FUNCTION_BLOCK fbShutterAct
VAR_INPUT
	Config :  stShutterConfig;
	OpenRelay : iRelay;
	CloseRelay : iRelay;
END_VAR
VAR_OUTPUT
	State : stShutterState;
END_VAR
VAR_IN_OUT

END_VAR
VAR
	CmdOpen : BOOL;
	CmdClose : BOOL;
	OutputCheckTimer : TON;
END_VAR

VAR CONSTANT
	OutputCheckCycleTime: TIME := T#50MS;
END_VAR
VAR RETAIN
	HeightTime: TIME := T#0S;
	AngleTime: TIME := T#0S;
END_VAR


// Both signals must not be set at the same time
IF CmdOpen AND CmdClose THEN
	CmdOpen := FALSE;
	CmdClose := FALSE;
END_IF

// Reset signal if shutter reached fully open position with overstep
IF CmdOpen AND HeightTime >= Config.HeightTravelTime + Config.HeightTravelTimeOverstep THEN
	CmdOpen := FALSE;
END_IF

// Reset signal if shutter reached fully close position
IF CmdClose AND HeightTime <= T#0S AND AngleTime <= T#0S THEN
	CmdClose := FALSE;
END_IF

// Write physical outputs and update shutter state
IF CmdOpen AND NOT CmdClose THEN
    CloseRelay.Reset();
    OpenRelay.Set();
	State.StateType := eShutterStateType.OPENING;
ELSIF CmdClose AND NOT CmdOpen THEN
    OpenRelay.Reset();
    CloseRelay.Set();
	State.StateType := eShutterStateType.CLOSING;
ELSE
    OpenRelay.Reset();
    CloseRelay.Reset();
	State.StateType := eShutterStateType.IDLE;
END_IF

// Count time and accumulate when signals are set
OutputCheckTimer(IN := CmdOpen OR CmdClose, PT := OutputCheckCycleTime);
IF OutputCheckTimer.Q THEN
	IF CmdOpen THEN
		// Open fins first before moving up
		IF AngleTime < Config.AngleTravelTime THEN
			AngleTime := AngleTime + OutputCheckCycleTime;
		ELSIF HeightTime < Config.HeightTravelTime THEN
			HeightTime := HeightTime + OutputCheckCycleTime;
		END_IF;
	END_IF
	
	IF CmdClose THEN
		// Close fins first before moving down
		IF AngleTime > T#0S THEN
			AngleTime := AngleTime - OutputCheckCycleTime;
		ELSIF HeightTime > T#0s THEN
			HeightTime := HeightTime - OutputCheckCycleTime;
		END_IF;
	END_IF
	
	OutputCheckTimer(IN := FALSE);  // reset
END_IF

// Update shutter position% basen on position time
State.Position.Height := TimeToPosition(CurrentPosTime := HeightTime, TravelTime := Config.HeightTravelTime);
State.Position.Angle := TimeToPosition(CurrentPosTime := AngleTime, TravelTime := Config.AngleTravelTime);

METHOD Close
CmdOpen := FALSE;
CmdClose := TRUE;
END_METHOD

METHOD Open
CmdClose := FALSE;
CmdOpen := TRUE;
END_METHOD

METHOD Stop
CmdOpen := FALSE;
CmdClose := FALSE;
END_METHOD

METHOD PUBLIC TimeToPosition : USINT
VAR_INPUT
	CurrentPosTime : TIME;
	TravelTime : TIME;
END_VAR
IF TravelTime <= T#0S THEN
    TimeToPosition := 0;
ELSE
    TimeToPosition := UDINT_TO_USINT(100 * TIME_TO_UDINT(CurrentPosTime) / TIME_TO_UDINT(TravelTime));
END_IF
END_METHOD

END_FUNCTION_BLOCK

(* stored: Version 1.1.0.1
   POU fbShutterAct: Id {1ba23f45-b0eb-421e-9a3b-6a879c5afe8f}, SpecialFunc None
   Method Close: Id {f613d1a9-dcd5-4ce8-bd35-546352718445}
   Method Open: Id {1dda91e8-cd15-4a31-9096-5e1a4c5f89a9}
   Method Stop: Id {17cc93a3-e742-4197-a775-db53f236a55d}
   Method TimeToPosition: Id {772cedc8-24ef-4e71-897a-f0415c3ffac2} *)
